// TIA Portal V16 export
FUNCTION "MCP_RC_FC5" : Void   // FC9805, LAD
{ S7_Optimized_Access := 'TRUE' }
   VAR_INPUT
      "a" : Bool;
   END_VAR
   VAR_OUTPUT
      q : Bool;
   END_VAR
BEGIN
END_FUNCTION
